INTERFACE I_Reversible EXTENDS I_Conveyor

PROPERTY Reverse : BOOL
GET
END_GET
SET
END_SET
END_PROPERTY

END_INTERFACE

(* stored: Version 1.1.0.1, ProductVersion 3.1 *)
